
// ===== library types =====

TYPE "UDT_Salidas_RFID"
   STRUCT
      Tag_escribir : Bool;   // Escribir en tag
      Tag_leer : Bool;   // Leer de tag
      Tag_reservado_2 : Bool;   // xBit2
      Tag_reservado_3 : Bool;   // xBit3
      Tag_antena_apagar : Bool;   // Apagar antena
      Tag_reservado_5 : Bool;   // xBit5
      Tag_reservado_6 : Bool;   // xBit6
      Tag_reservado_7 : Bool;   // xBit7
      Reservado_AB5 : Byte;   // byReserved
      Tag_direccion_leer_escribir : Word;   // Direccion de R/W
      Tag_datos_a_escribir : Array[0..27] of Byte;   // Datos a escribir
   END_STRUCT;
END_TYPE

TYPE "UDT_Estado"
   STRUCT
      Modo_auto : Bool;   // Marca Modo
      Modo_manual : Bool;   // Marca Modo
      Ciclo_auto_activo : Bool;   // Marca Modo
      Ciclo_manual_activo : Bool;   // Marca Modo
      Emergencia : Bool;   // Marca Modo
      Rearme_requerido : Bool;   // Marca Modo
      Marcha_permitida : Bool;   // Marca Modo
      Condicion_arranque_auto : Bool;   // Marca Condiciones
      Condicion_arranque_manual : Bool;   // Marca Condiciones
      Estacion_cond_iniciales : Bool;   // Marca Condiciones
      Cinta_habilitada : Bool;   // Marca Condiciones
      Ciclo_manual_terminado : Bool;   // Marca Condiciones
      Rearme_requerido_gestion : Bool;   // Marca Condiciones
      Palet_en_posicion : Bool;   // Marca Cinta
      Palet_en_estacion : Bool;   // Marca Cinta
      Palet_evacuado : Bool;   // Marca Cinta
      Orden_evacuar : Bool;   // Marca Cinta
      Orden_leer : Bool;   // Marca RFID
      Orden_escribir : Bool;   // Marca RFID
      Rfid_lectura_ok : Bool;   // Marca RFID
      Rfid_escritura_ok : Bool;   // Marca RFID
      Rfid_error : Bool;   // Marca RFID
      Rfid_codigo_error : Byte;   // Marca RFID
      App_inicio : Bool;   // Marca App
      App_en_reposo : Bool;   // Marca App
      App_terminada : Bool;   // Marca App
      App_alarma : Bool;
   END_STRUCT;
END_TYPE

TYPE "UDT_Entradas_Basico"
   STRUCT
      Boton_marcha : Bool;   // Botón de marcha
      Boton_paro : Bool;   // Botón de paro (0 activado)
      Selector_modo : Bool;   // Selector Manual/Auto (0 - Manual / 1 - Auto)
      Boton_rearme : Bool;   // Botón de rearme
      Sensor_ind_bien_pos : Bool;   // Palet bien posicionado - Sensor inductivo 0 (Extremo derecho)
      Seta_emergencia : Bool;   // Seta de emergencia
      Sensor_palet_izq : Bool;   // Palet en extremo izquierdo
      Sensor_palet_dch : Bool;   // Palet en extremo derecho
   END_STRUCT;
END_TYPE

TYPE "UDT_Entradas_Stopper"
   STRUCT
      Sensor_ind_0 : Bool;   // Entrada Sensor inductivo 0 (Extremo derecho)
      Sensor_ind_1 : Bool;   // Entrada Sensor inductivo 1
      Sensor_ind_2 : Bool;   // Entrada Sensor inductivo 2
      Sensor_ind_3 : Bool;   // Entrada Sensor inductivo 3 (Extremo izquierdo)
      Reservado_E2_4 : Bool;
      Reservado_E2_5 : Bool;
      Reservado_E2_6 : Bool;
      Sensor_stopper_abajo : Bool;   // Entrada Stopper abajo
   END_STRUCT;
END_TYPE

TYPE "UDT_Salidas_Basico"
   STRUCT
      Led_boton_marcha : Bool;   // Luz del boton de Marcha
      Led_boton_rearme : Bool;   // Luz del boton de Reset
      Led_q1_ciclo_auto : Bool;   // Luz Q1
      Led_q2_emergencia : Bool;   // Luz Q2
      Cinta_dch : Bool;   // Arrancar cinta hacia la derecha
      Cinta_izq : Bool;   // Arrancar cinta hacia la izquierda
      Cinta_velocidad_baja : Bool;   // Establecer velocidad baja
      Bajar_stopper : Bool;   // Bajar cilindro Stopper
   END_STRUCT;
END_TYPE

TYPE "UDT_Entradas_RFID"
   STRUCT
      Tag_datos_escritos : Bool;   // Datos escritos
      Tag_datos_leidos : Bool;   // Datos leidos
      Reservado_E4_2 : Bool;
      Reservado_E4_3 : Bool;
      Tag_antena_apagada : Bool;   // Antena apagada
      Tag_detectado : Bool;   // Tag detectado
      Tag_error : Bool;   // Error
      Tag_proceso_listo : Bool;   // Proceso listo
      Tag_codigo_error : Byte;   // Codigo de error
      Tag_direccion_confirmada : Word;   // Direccion de escritura
      Tag_datos_leidos_escritos : Array[0..27] of Byte;   // Datos
   END_STRUCT;
END_TYPE

FUNCTION_BLOCK "Est_FB_Estacion"   // FB1, SCL
{ S7_Optimized_Access := 'TRUE' }
VERSION : 0.1
   VAR_INPUT
      InBasico : "UDT_Entradas_Basico";
      InRFID : "UDT_Entradas_RFID";
      InStopper : "UDT_Entradas_Stopper";
      Direccion_lectura : Word;
      Direccion_escritura : Word;
      App_en_reposo : Bool;
      App_terminada : Bool;
      App_alarma : Bool;
      App_rearme_requerido : Bool;
      Inhibir_cinta : Bool;
      Mascara_lectura : DWord := 16#0FFFFFFF;
      Mascara_escritura : DWord;
   END_VAR
   VAR_OUTPUT
      App_inicio : Bool;
      Emergencia : Bool;
      Rearme : Bool;
   END_VAR
   VAR_IN_OUT
      OutBasico : "UDT_Salidas_Basico";
      OutRFID : "UDT_Salidas_RFID";
      Imagen_palet : Array[0..27] of Byte;
   END_VAR
   VAR
      Etapa_gestion : Int;
      Etapa_0 : Bool;
      Etapa_1 : Bool;
      Etapa_2 : Bool;
      Etapa_3 : Bool;
      Etapa_4 : Bool;
      Etapa_5 : Bool;
      Estado_Estacion : "UDT_Estado";
      Flanco_rearme : R_TRIG;
      FB2_Modo_Instance : "Est_FB_Modo";
      FB3_Cinta_Instance : "Est_FB_Cinta";
      FB4_RFID_Instance : "Est_FB_RFID";
      Ciclo_manual_acabado : Bool;
   END_VAR
BEGIN
   #Estado_Estacion.App_en_reposo := #App_en_reposo;
   #Estado_Estacion.App_terminada := #App_terminada;
   #Estado_Estacion.App_alarma := #App_alarma;

   //Flanco de rearme
   #Flanco_rearme(CLK := #InBasico.Boton_rearme);

   //Condiciones combinacionales
   //las CI han cambiado ahora que tenemos app
   // Tensión en la máquina (24 Vdc) – No existe señal de PLC.
   // Aire comprimido (6 bar) – No existe señal de PLC.
   // Debe existir un palet correctamente posicionado.
   // El cilindro eje vertical Debe estar en su posición extrema superior.
   // El cilindro eje horizontal Debe estar referenciado.
   // La garra estará en posición de reposo (desctivada/cerrada).
   // No existe estado de emergencia.
   #Estado_Estacion.Estacion_cond_iniciales := NOT #Estado_Estacion.Emergencia AND NOT #InStopper.Sensor_stopper_abajo AND #Estado_Estacion.App_en_reposo
   AND NOT #Estado_Estacion.Rfid_error;

   #Estado_Estacion.Condicion_arranque_auto := #Estado_Estacion.Estacion_cond_iniciales;
   #Estado_Estacion.Condicion_arranque_manual := #Estado_Estacion.Estacion_cond_iniciales AND #Estado_Estacion.Palet_en_estacion;

   #Estado_Estacion.Cinta_habilitada := (#Estado_Estacion.Ciclo_auto_activo OR #Estado_Estacion.Ciclo_manual_activo) AND NOT #Estado_Estacion.Emergencia;

   //llamo a Modo
   #FB2_Modo_Instance(Seta_emergencia := NOT #InBasico.Seta_emergencia,
                      Boton_rearme := #InBasico.Boton_rearme,
                      Boton_marcha := #InBasico.Boton_marcha,
                      Boton_paro := NOT #InBasico.Boton_paro,
                      Selector_automatico := #InBasico.Selector_modo,
                      Condicion_arranque_auto := #Estado_Estacion.Condicion_arranque_auto,
                      Condicion_arranque_manual := #Estado_Estacion.Condicion_arranque_manual,
                      Ciclo_manual_acabado := #Ciclo_manual_acabado,
                      Modo_auto := #Estado_Estacion.Modo_auto,
                      Modo_manual := #Estado_Estacion.Modo_manual,
                      Ciclo_auto_activo := #Estado_Estacion.Ciclo_auto_activo,
                      Ciclo_manual_activo := #Estado_Estacion.Ciclo_manual_activo,
                      Emergencia := #Estado_Estacion.Emergencia,
                      Rearme_requerido := #Estado_Estacion.Rearme_requerido,
                      Marcha_permitida := #Estado_Estacion.Marcha_permitida
   );

   //gestión
   CASE #Etapa_gestion OF
       0:  // ESPERA PALET
           IF (#Estado_Estacion.Ciclo_auto_activo OR #Estado_Estacion.Ciclo_manual_activo) AND #Estado_Estacion.Palet_en_posicion AND NOT #Estado_Estacion.Emergencia THEN
               #Etapa_gestion := 1;
           END_IF;
       1:  // LEER RFID
           IF #Estado_Estacion.Rfid_error THEN
               #Etapa_gestion := 6;
           ELSIF #Estado_Estacion.Rfid_lectura_ok THEN
               #Etapa_gestion := 2;
           END_IF;
       2:  // APLICACION
           IF #Estado_Estacion.App_terminada THEN
               #Etapa_gestion := 3;
           END_IF;
       3:  // ESCRIBIR RFID
           IF #Estado_Estacion.Rfid_error THEN
               #Etapa_gestion := 6;
           ELSIF #Estado_Estacion.Rfid_escritura_ok THEN
               #Etapa_gestion := 4;
           END_IF;
       4:  // EVACUAR
           IF #Estado_Estacion.Palet_evacuado THEN
               #Etapa_gestion := 5;
           END_IF;
       5:  // FIN PALET
           #Etapa_gestion := 0;
       6:  // FALLO RFID
           IF #Flanco_rearme.Q THEN
               #Etapa_gestion := 4;
           END_IF;
       ELSE
           #Etapa_gestion := 0;
   END_CASE;

   //Emergencia
   IF #Estado_Estacion.Emergencia THEN
       #Etapa_gestion := 0;
   END_IF;

   //Ordenes
   #Estado_Estacion.Orden_leer := (#Etapa_gestion = 1);
   #Estado_Estacion.App_inicio := (#Etapa_gestion = 2);
   #Estado_Estacion.Orden_escribir := (#Etapa_gestion = 3);
   #Estado_Estacion.Orden_evacuar := (#Etapa_gestion = 4);
   #Ciclo_manual_acabado := (#Etapa_gestion = 5 OR (#Etapa_gestion = 0 AND NOT #Estado_Estacion.Palet_en_estacion))
   AND #Estado_Estacion.Modo_manual;
   #Estado_Estacion.Rearme_requerido_gestion := (#Etapa_gestion = 6);

   //Cadenas
   #FB3_Cinta_Instance(Cinta_habilitada := #Estado_Estacion.Cinta_habilitada,
                       Orden_evacuar := #Estado_Estacion.Orden_evacuar,
                       Emergencia := #Estado_Estacion.Emergencia,
                       Sensor_palet_izq := #InBasico.Sensor_palet_izq,
                       Sensor_palet_dch := #InBasico.Sensor_palet_dch,
                       Sensor_ind_bien_pos := #InBasico.Sensor_ind_bien_pos,
                       Sensor_stopper_abajo := #InStopper.Sensor_stopper_abajo,
                       Cinta_dch := #OutBasico.Cinta_dch,
                       Bajar_stopper := #OutBasico.Bajar_stopper,
                       Palet_en_posicion := #Estado_Estacion.Palet_en_posicion,
                       Palet_en_estacion := #Estado_Estacion.Palet_en_estacion,
                       Palet_evacuado := #Estado_Estacion.Palet_evacuado
   );

   IF #Inhibir_cinta THEN
       #OutBasico.Cinta_dch := FALSE;
   END_IF;

   #FB4_RFID_Instance(Orden_leer := #Estado_Estacion.Orden_leer,
                      Orden_escribir := #Estado_Estacion.Orden_escribir,
                      Emergencia := #Estado_Estacion.Emergencia,
                      Tag_datos_escritos := #InRFID.Tag_datos_escritos,
                      Tag_datos_leidos := #InRFID.Tag_datos_leidos,
                      Tag_antena_apagada := #InRFID.Tag_antena_apagada,
                      Tag_detectado := #InRFID.Tag_detectado,
                      Tag_error := #InRFID.Tag_error,
                      Tag_proceso_listo := #InRFID.Tag_proceso_listo,
                      Tag_codigo_error := #InRFID.Tag_codigo_error,
                      Tag_direccion_confirmada := #InRFID.Tag_direccion_confirmada,
                      Tag_datos_leidos_escritos := #InRFID.Tag_datos_leidos_escritos,
                      Mascara_lectura:=#Mascara_lectura,
                      Mascara_escritura:=#Mascara_escritura,
                      Tag_escribir := #OutRFID.Tag_escribir,
                      Tag_leer := #OutRFID.Tag_leer,
                      Tag_antena_apagar := #OutRFID.Tag_antena_apagar,
                      Tag_direccion_leer_escribir := #OutRFID.Tag_direccion_leer_escribir,
                      Tag_datos_a_escribir := #OutRFID.Tag_datos_a_escribir,
                      Rfid_lectura_ok := #Estado_Estacion.Rfid_lectura_ok,
                      Rfid_escritura_ok := #Estado_Estacion.Rfid_escritura_ok,
                      Rfid_error := #Estado_Estacion.Rfid_error,
                      Rfid_codigo_error := #Estado_Estacion.Rfid_codigo_error,
                      Imagen:=#Imagen_palet,
                      Direccion_escritura:=#Direccion_escritura,
                      Direccion_lectura:=#Direccion_lectura);

   #App_inicio := #Estado_Estacion.App_inicio;
   #Emergencia := #Estado_Estacion.Emergencia;
   #Rearme := #Flanco_rearme.Q;

   //Luces del panel y salidas sin uso
   #OutBasico.Led_boton_marcha := #Estado_Estacion.Marcha_permitida;
   #OutBasico.Led_boton_rearme := #Estado_Estacion.Rearme_requerido OR #Estado_Estacion.Rearme_requerido_gestion OR #App_rearme_requerido;
   #OutBasico.Led_q1_ciclo_auto := #Estado_Estacion.Ciclo_auto_activo;
   #OutBasico.Led_q2_emergencia := #Estado_Estacion.Emergencia OR (#Estado_Estacion.App_alarma);// AND "Clock_1Hz");
   #OutBasico.Cinta_izq := FALSE;
   #OutBasico.Cinta_velocidad_baja := FALSE;
END_FUNCTION_BLOCK

FUNCTION_BLOCK "Est_FB_Modo"   // FB2, SCL
{ S7_Optimized_Access := 'TRUE' }
VERSION : 0.1
   VAR_INPUT
      Seta_emergencia : Bool;
      Boton_rearme : Bool;
      Boton_marcha : Bool;
      Boton_paro : Bool;
      Selector_automatico : Bool;
      Condicion_arranque_auto : Bool;
      Condicion_arranque_manual : Bool;
      Ciclo_manual_acabado : Bool;
   END_VAR
   VAR_IN_OUT
      Modo_auto : Bool;
      Modo_manual : Bool;
      Ciclo_auto_activo : Bool;
      Ciclo_manual_activo : Bool;
      Emergencia : Bool;
      Rearme_requerido : Bool;
      Marcha_permitida : Bool;
   END_VAR
   VAR
      Etapa_emergencia : Int := 10;
      Etapa_modo : Int := 20;
      Etapa_ciclo : Int := 30;
      Flanco_marcha : R_TRIG;
      Flanco_rearme : R_TRIG;
   END_VAR
BEGIN
   #Modo_auto := FALSE;
   #Modo_manual := FALSE;
   #Ciclo_auto_activo := FALSE;
   #Ciclo_manual_activo := FALSE;
   #Emergencia := FALSE;
   #Rearme_requerido := FALSE;
   #Marcha_permitida := FALSE;

   #Flanco_marcha(CLK:=#Boton_marcha);
   #Flanco_rearme(CLK:=#Boton_rearme);

   CASE #Etapa_emergencia OF
       10:  //NORMAL
           IF #Seta_emergencia THEN
               #Etapa_emergencia := 11;
           END_IF;
           ;
       11:  //EMERGENCIA
           #Emergencia := TRUE;
           #Rearme_requerido := TRUE;
           IF #Flanco_rearme.Q AND NOT #Seta_emergencia THEN
               #Etapa_emergencia := 10;
           END_IF;
           ;
       ELSE
           #Etapa_emergencia := 11;
           ;
   END_CASE;

   CASE #Etapa_modo OF
       20:  // MANUAL
           #Modo_manual := TRUE;
           IF #Selector_automatico THEN
               #Etapa_modo := 21;
           END_IF;
           ;
       21:  // AUTOMATICO
           #Modo_auto := TRUE;
           IF NOT #Selector_automatico THEN
               #Etapa_modo := 20;
           END_IF;
           ;
       ELSE
           #Etapa_modo := 20;
           #Etapa_emergencia := 11;
           ;
   END_CASE;

   CASE #Etapa_ciclo OF
       30:  // REPOSO
           IF NOT #Emergencia AND ((#Modo_auto AND #Condicion_arranque_auto) OR (#Modo_manual AND #Condicion_arranque_manual)) THEN
               #Marcha_permitida := TRUE;
           END_IF;

           IF #Marcha_permitida AND #Flanco_marcha.Q AND #Modo_auto THEN
               #Etapa_ciclo := 31;
           ELSIF #Marcha_permitida AND #Flanco_marcha.Q AND #Modo_manual THEN
               #Etapa_ciclo := 32;
           END_IF;
           ;
       31:  // AUTOMATICO ACTIVO
           #Ciclo_auto_activo := TRUE;
           IF #Boton_paro OR #Emergencia OR NOT #Modo_auto THEN
               #Etapa_ciclo := 30;
           END_IF;
           ;
       32:  //MANUAL ACTIVO
           #Ciclo_manual_activo := TRUE;
           IF #Boton_paro OR #Emergencia OR NOT #Modo_manual OR #Ciclo_manual_acabado THEN
               #Etapa_ciclo := 30;
           END_IF;
           ;
       ELSE
           #Etapa_ciclo := 30;
           #Etapa_emergencia := 11;
           ;
   END_CASE;
END_FUNCTION_BLOCK

FUNCTION_BLOCK "Est_FB_Cinta"   // FB3, SCL
{ S7_Optimized_Access := 'TRUE' }
VERSION : 0.1
   VAR_INPUT
      Emergencia : Bool;   // De modo
      Cinta_habilitada : Bool;   // ciclo activo y estación en condiciones iniciales
      Orden_evacuar : Bool;   // la aplicación ya terminó y el RFID está escrito
      Sensor_palet_izq : Bool;   // Extremos de la cinta
      Sensor_palet_dch : Bool;   // Extremos de la cinta
      Sensor_ind_bien_pos : Bool;   // Palet apoyado en el stopper
      Sensor_stopper_abajo : Bool;   // Confirmación del stopper
   END_VAR
   VAR_IN_OUT
      Cinta_dch : Bool;   // Actuadores
      Bajar_stopper : Bool;   // Actuadores
      Palet_en_posicion : Bool;   // Hay palet listo para trabajar
      Palet_en_estacion : Bool;   // Sensor_palet_izq + Sensor_palet_dch + Sensor_ind_bien_pos, para Condicion_arranque_manual
      Palet_evacuado : Bool;   // activa Ciclo_manual_terminado
   END_VAR
   VAR
      Etapa_cinta : Int;   // nuemero de etapa
      Etapa_2 : Bool;   // estamos en la 2
      Timer_etapa2 : TON_TIME;   // timer de la 2
      Flanco_subida_sensor_palet_dch : R_TRIG;   // flanco subida del sensor
      Flanco_bajada_sensor_palet_dch : F_TRIG;   // flanco bajada del sensor
      Palets_en_cinta : Int;
      Flanco_subida_sensor_palet_izq : R_TRIG;
      Timer_Stopper_Etapa5 : TON_TIME;
      Timer_avance : TON_TIME;
   END_VAR
BEGIN

   #Cinta_dch := FALSE;
   #Palet_en_posicion := FALSE;
   #Palet_en_estacion := FALSE;
   #Etapa_2 := FALSE;
   #Palet_evacuado := FALSE;

   #Flanco_subida_sensor_palet_dch(CLK := #Sensor_palet_dch);
   #Flanco_bajada_sensor_palet_dch(CLK := #Sensor_palet_dch);
   #Flanco_subida_sensor_palet_izq(CLK := #Sensor_palet_izq);
   #Timer_Stopper_Etapa5(IN := #Etapa_cinta = 5,
                         PT := T#400ms);
   #Timer_avance(IN := #Etapa_cinta = 1 OR #Etapa_cinta = 6, PT := T#10s);



   IF #Etapa_cinta = 2 THEN
       #Etapa_2 := TRUE;
   END_IF;

   #Timer_etapa2(IN := #Etapa_2,
                 PT := T#300ms);

   IF #Flanco_subida_sensor_palet_izq.Q THEN
       #Palets_en_cinta := #Palets_en_cinta + 1;
   END_IF;
   IF #Flanco_bajada_sensor_palet_dch.Q AND #Palets_en_cinta > 0 THEN
       #Palets_en_cinta := #Palets_en_cinta - 1;
   END_IF;

   IF #Sensor_ind_bien_pos AND #Palets_en_cinta = 0 THEN
       #Palets_en_cinta := 1;
   END_IF;

   CASE #Etapa_cinta OF
       0:  // PARADA
           #Cinta_dch := FALSE;
           #Bajar_stopper := FALSE;
           IF #Cinta_habilitada AND (#Sensor_palet_izq OR #Palets_en_cinta > 0) AND NOT #Sensor_ind_bien_pos THEN
               #Etapa_cinta := 1;
           ELSIF #Cinta_habilitada AND #Sensor_ind_bien_pos THEN
               #Etapa_cinta := 3;
           END_IF;
       1:  //AVANCE
           #Cinta_dch := TRUE;
           IF #Sensor_ind_bien_pos THEN
               #Etapa_cinta := 3;
           ELSIF #Timer_avance.Q THEN   // no llega ningun palet: el contador estaba descuadrado
               #Palets_en_cinta := 0;
               #Etapa_cinta := 0;
           END_IF;
       2:  //ASENTAR
           #Cinta_dch := TRUE;
           IF #Timer_etapa2.Q THEN
               #Etapa_cinta := 3;
           END_IF;
       3:  //PALET EN POSICION
           #Palet_en_posicion := TRUE;
           IF #Orden_evacuar THEN
               #Etapa_cinta := 4;
           END_IF;
       4:  //LIBERAR
           #Bajar_stopper := TRUE;
           IF NOT #Sensor_stopper_abajo THEN
               #Etapa_cinta := 5;
           END_IF;
       5:  //SACAR
           #Bajar_stopper := TRUE;
           #Cinta_dch := TRUE;
           IF #Timer_Stopper_Etapa5.Q OR #Flanco_subida_sensor_palet_dch.Q THEN
               #Etapa_cinta := 6;
               ;
           END_IF;
       6: //SALIR
           #Bajar_stopper := FALSE;
           #Cinta_dch := TRUE;
           IF #Flanco_bajada_sensor_palet_dch.Q THEN
               #Etapa_cinta := 7;
               ;
           ELSIF #Timer_avance.Q THEN   // el palet no pasa por el sensor (retirado a mano): no dejar la cinta en marcha
               #Palets_en_cinta := 0;
               #Etapa_cinta := 7;
           END_IF;
       7: //TERMINAR
           #Palet_evacuado := TRUE;
           #Etapa_cinta := 0;
       ELSE  // Statement section ELSE
           #Etapa_cinta := 0;
           ;
   END_CASE;

   #Palet_en_estacion := #Sensor_palet_dch OR #Sensor_palet_izq OR #Sensor_ind_bien_pos OR (#Palets_en_cinta > 0) OR #Etapa_cinta = 1;

   IF #Emergencia THEN
       #Etapa_cinta := 0;
       #Cinta_dch := FALSE;
       #Bajar_stopper := FALSE;
       #Palets_en_cinta := 0;   // el operario retira los palets en la emergencia
   END_IF;
END_FUNCTION_BLOCK

FUNCTION_BLOCK "Est_FB_RFID"   // FB4, SCL
{ S7_Optimized_Access := 'TRUE' }
VERSION : 0.1
   VAR_INPUT
      Emergencia : Bool;
      Orden_escribir : Bool;
      Orden_leer : Bool;
      Tag_datos_escritos : Bool;
      Tag_datos_leidos : Bool;
      Tag_antena_apagada : Bool;
      Tag_detectado : Bool;
      Tag_error : Bool;
      Tag_proceso_listo : Bool;
      Tag_codigo_error : Byte;
      Tag_direccion_confirmada : Word;
      Tag_datos_leidos_escritos : Array[0..27] of Byte;
      Direccion_lectura : Word;
      Direccion_escritura : Word;
      Mascara_lectura : DWord;
      Mascara_escritura : DWord;
   END_VAR
   VAR_IN_OUT
      Tag_escribir : Bool;
      Tag_leer : Bool;
      Tag_antena_apagar : Bool;
      Tag_direccion_leer_escribir : Word;
      Tag_datos_a_escribir : Array[0..27] of Byte;
      Rfid_lectura_ok : Bool;
      Rfid_escritura_ok : Bool;
      Rfid_error : Bool;
      Rfid_codigo_error : Byte;
      Imagen : Array[0..27] of Byte;
   END_VAR
   VAR
      T_Rfid : TON_TIME;
      Etapa_rfid : Int;
      Etapa_1 : Bool;
      Etapa_3 : Bool;
      Etapa_4 : Bool;
      Rfid_ocupado : Bool;
      Imagen_leida : Array[0..27] of Byte;
   END_VAR
   VAR_TEMP
      i : Int;
   END_VAR
BEGIN
   //PARA EL DANI DEL FUTURO
   //que vaya leyendo los codigos rfid por si me vienen dos palets juntos
   //y que los meta en una cola para luego leerlos y escribirlos por orden?
   //      - no lo voy a hacer porque creo que esto solo es un problema en el simulador
   //      - pero gracias por la idea dani del pasado
   //---------------------------------------------------------------------------
   #Tag_escribir := FALSE;
   #Tag_leer := FALSE;
   #Tag_antena_apagar := TRUE;
   #Rfid_lectura_ok := FALSE;
   #Rfid_escritura_ok := FALSE;
   #Rfid_error := FALSE;
   #Etapa_1 := FALSE;
   #Etapa_3 := FALSE;
   #Etapa_4 := FALSE;

   CASE #Etapa_rfid OF
       0:  // REPOSO
           #Tag_antena_apagar := TRUE;
           #Tag_leer := FALSE;
           #Tag_escribir := FALSE;
           IF (#Orden_leer OR #Orden_escribir) AND NOT #Emergencia THEN
               #Etapa_rfid := 1;
               ;
           END_IF;
       1:  // ENERGIZAR
           #Tag_antena_apagar := FALSE;
           #Etapa_1 := TRUE;
           IF #Tag_error OR #T_Rfid.Q THEN
               #Etapa_rfid := 8;
           ELSIF NOT #Tag_antena_apagada AND #Tag_detectado AND #Tag_proceso_listo AND NOT #Tag_error THEN
               #Etapa_rfid := 2;
           END_IF;
           ;
       2:  // LISTO
           #Tag_antena_apagar := FALSE;
           #Rfid_ocupado := FALSE;
           IF #Orden_leer AND NOT #Orden_escribir THEN
               #Etapa_rfid := 3;
           ELSIF NOT #Orden_leer AND #Orden_escribir THEN
               #Etapa_rfid := 4;
           END_IF;
           ;
       3:  // LEER
           #Tag_antena_apagar := FALSE;
           #Etapa_3 := TRUE;
           // "leido" es el eco de la orden: el dato solo vale cuando "listo" baja y vuelve a subir
           IF NOT #Tag_proceso_listo THEN
               #Rfid_ocupado := TRUE;
           END_IF;
           #Tag_leer := TRUE;
           #Tag_direccion_leer_escribir := #Direccion_lectura;
           IF #Tag_error OR #T_Rfid.Q THEN
               #Etapa_rfid := 8;
           ELSIF #Rfid_ocupado AND #Tag_datos_leidos AND #Tag_proceso_listo AND #Tag_direccion_confirmada = #Direccion_lectura THEN
               #Imagen_leida := #Tag_datos_leidos_escritos;   // copia completa se usa al escribir
               FOR #i := 0 TO 27 DO
                   IF (SHR(IN := #Mascara_lectura, N := #i) AND 16#1) <> 16#0 THEN
                       #Imagen[#i] := #Tag_datos_leidos_escritos[#i];
                   ELSE
                       #Imagen[#i] := 0;   // lo que no es de esta estacion no pasa a la app
                   END_IF;
               END_FOR;
               #Etapa_rfid := 5;
           END_IF;
           ;
       4:  // ESCRIBIR
           #Tag_antena_apagar := FALSE;
           #Etapa_4 := TRUE;
           IF NOT #Tag_proceso_listo THEN
               #Rfid_ocupado := TRUE;
           END_IF;
           #Tag_escribir := TRUE;
           #Tag_direccion_leer_escribir := #Direccion_escritura;
           FOR #i := 0 TO 27 DO
               IF (SHR(IN := #Mascara_escritura, N := #i) AND 16#1) <> 16#0 THEN
                   #Tag_datos_a_escribir[#i] := #Imagen[#i];       // byte de esta estacion
               ELSE
                   #Tag_datos_a_escribir[#i] := #Imagen_leida[#i]; // byte ajeno: se devuelve como estaba
               END_IF;
           END_FOR;
           IF #Tag_error OR #T_Rfid.Q THEN
               #Etapa_rfid := 8;
           ELSIF #Rfid_ocupado AND #Tag_datos_escritos AND #Tag_proceso_listo AND #Tag_direccion_confirmada = #Direccion_escritura THEN
               #Etapa_rfid := 6;
           END_IF;
           ;
       5:  // LEIDO
           #Tag_antena_apagar := FALSE;
           #Rfid_lectura_ok := TRUE;
           IF NOT #Orden_leer THEN
               #Etapa_rfid := 0;
           END_IF;
           ;
       6:  // ESCRITO 
           #Tag_antena_apagar := FALSE;
           #Rfid_escritura_ok := TRUE;
           IF NOT #Orden_escribir THEN
               #Etapa_rfid := 0;
           END_IF;
           ;
       8:  // ERROR RFID
           #Rfid_error := TRUE;
           #Rfid_codigo_error := #Tag_codigo_error;
           #Tag_antena_apagar := TRUE;
           #Tag_leer := FALSE;
           #Tag_escribir := FALSE;
           IF NOT #Orden_escribir AND NOT #Orden_leer THEN   // CIROS no da "antena apagada" (iAntenaOFF sin conectar)
               #Etapa_rfid := 0;
           END_IF;
           ;
       ELSE  // Statement section ELSE
           #Etapa_rfid := 0;
           ;
   END_CASE;

   #T_Rfid(IN := #Etapa_1 OR #Etapa_3 OR #Etapa_4,
           PT := T#5s);

   IF #Emergencia THEN
       #Etapa_rfid := 0;
       #Tag_antena_apagar := TRUE;
       #Tag_escribir := FALSE;
       #Tag_leer := FALSE;
       #Rfid_lectura_ok := FALSE;
       #Rfid_escritura_ok := FALSE;
       #Rfid_error := FALSE;
   END_IF;
END_FUNCTION_BLOCK

// ===== library: MasterCopy "Main" =====

ORGANIZATION_BLOCK "Main"   // OB1, LAD, ProgramCycle
TITLE = "Main Program Sweep (Cycle)"
{ S7_Optimized_Access := 'TRUE' }
VERSION : 0.1
   VAR_INPUT
      Initial_Call : Bool;   // Initial call of this OB
      Remanence : Bool;   // =True, if remanent data are available
   END_VAR
BEGIN

REGION Network 1: Llamada al gestor
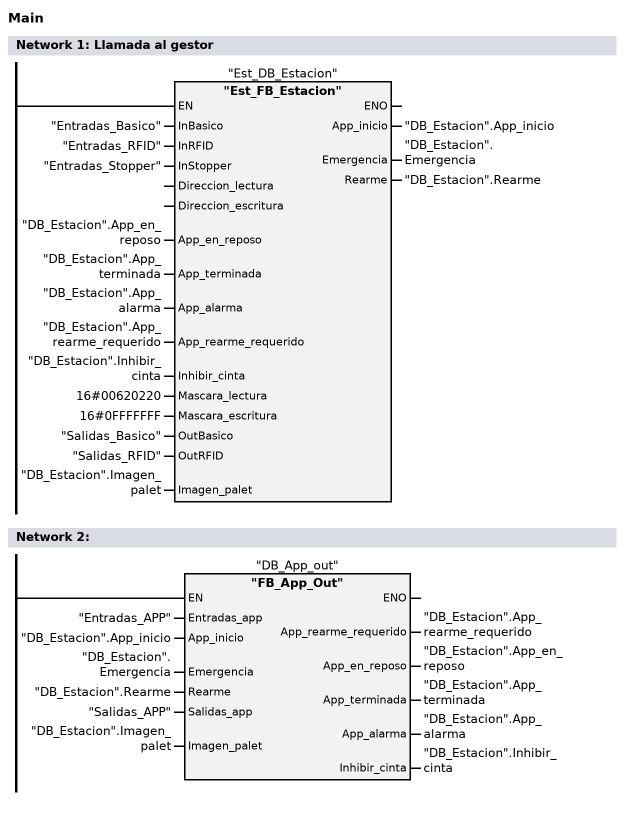
   RUNG wire#powerrail
      "Est_DB_Estacion"(InBasico := "Entradas_Basico", InRFID := "Entradas_RFID", InStopper := "Entradas_Stopper", Direccion_lectura :=, Direccion_escritura :=, App_en_reposo := "DB_Estacion".App_en_reposo, App_terminada := "DB_Estacion".App_terminada, App_alarma := "DB_Estacion".App_alarma, App_rearme_requerido := "DB_Estacion".App_rearme_requerido, Inhibir_cinta := "DB_Estacion".Inhibir_cinta, Mascara_lectura := 16#00620220, Mascara_escritura := 16#0FFFFFFF, OutBasico := "Salidas_Basico", OutRFID := "Salidas_RFID", Imagen_palet := "DB_Estacion".Imagen_palet, App_inicio => "DB_Estacion".App_inicio, Emergencia => "DB_Estacion".Emergencia, Rearme => "DB_Estacion".Rearme)
   END_RUNG
   // the same network as SCL:
   "Est_DB_Estacion"(InBasico := "Entradas_Basico",   // "Est_FB_Estacion"
                     InRFID := "Entradas_RFID",
                     InStopper := "Entradas_Stopper",
                     App_en_reposo := "DB_Estacion".App_en_reposo,
                     App_terminada := "DB_Estacion".App_terminada,
                     App_alarma := "DB_Estacion".App_alarma,
                     App_rearme_requerido := "DB_Estacion".App_rearme_requerido,
                     Inhibir_cinta := "DB_Estacion".Inhibir_cinta,
                     Mascara_lectura := 16#00620220,
                     Mascara_escritura := 16#0FFFFFFF,
                     OutBasico := "Salidas_Basico",
                     OutRFID := "Salidas_RFID",
                     Imagen_palet := "DB_Estacion".Imagen_palet,
                     App_inicio => "DB_Estacion".App_inicio,
                     Emergencia => "DB_Estacion".Emergencia,
                     Rearme => "DB_Estacion".Rearme);
END_REGION

REGION Network 2
   RUNG wire#powerrail
      "DB_App_out"(Entradas_app := "Entradas_APP", App_inicio := "DB_Estacion".App_inicio, Emergencia := "DB_Estacion".Emergencia, Rearme := "DB_Estacion".Rearme, Salidas_app := "Salidas_APP", Imagen_palet := "DB_Estacion".Imagen_palet, App_rearme_requerido => "DB_Estacion".App_rearme_requerido, App_en_reposo => "DB_Estacion".App_en_reposo, App_terminada => "DB_Estacion".App_terminada, App_alarma => "DB_Estacion".App_alarma, Inhibir_cinta => "DB_Estacion".Inhibir_cinta)
   END_RUNG
   // the same network as SCL:
   "DB_App_out"(Entradas_app := "Entradas_APP",   // "FB_App_Out"
                App_inicio := "DB_Estacion".App_inicio,
                Emergencia := "DB_Estacion".Emergencia,
                Rearme := "DB_Estacion".Rearme,
                Salidas_app := "Salidas_APP",
                Imagen_palet := "DB_Estacion".Imagen_palet,
                App_rearme_requerido => "DB_Estacion".App_rearme_requerido,
                App_en_reposo => "DB_Estacion".App_en_reposo,
                App_terminada => "DB_Estacion".App_terminada,
                App_alarma => "DB_Estacion".App_alarma,
                Inhibir_cinta => "DB_Estacion".Inhibir_cinta);
END_REGION
END_ORGANIZATION_BLOCK

// ===== library: MasterCopy "DB_Estacion" =====

DATA_BLOCK "DB_Estacion"   // DB2
{ S7_Optimized_Access := 'TRUE' }
VERSION : 0.1
   VAR
      Imagen_palet : Array[0..27] of Byte;
      App_inicio : Bool;
      App_en_reposo : Bool;
      App_terminada : Bool;
      App_alarma : Bool;
      App_rearme_requerido : Bool;
      Inhibir_cinta : Bool;
      Emergencia : Bool;
      Rearme : Bool;
   END_VAR
BEGIN
END_DATA_BLOCK

// ===== library: MasterCopy "FB_App_Out" =====

FUNCTION_BLOCK "FB_App_Out"   // FB5, SCL
{ S7_Optimized_Access := 'TRUE' }
VERSION : 0.1
   VAR_INPUT
      Entradas_app : "UDT_Entradas_APP";
      App_inicio : Bool;
      Emergencia : Bool;
      Rearme : Bool;
   END_VAR
   VAR_OUTPUT
      App_rearme_requerido : Bool;
      App_en_reposo : Bool;
      App_terminada : Bool;
      App_alarma : Bool;
      Inhibir_cinta : Bool;
   END_VAR
   VAR_IN_OUT
      Salidas_app : "UDT_Salidas_APP";
      Imagen_palet : Array[0..27] of Byte;
   END_VAR
   VAR
      Cond_conf : Bool;
      Cond_almacen : Bool;
      Etapa_app : Int;
      Etapa_previa : Int;
      Posicion_objetivo : Int;
      Almacen_destino : Int;
      Start_enviado : Bool;
      Pieza_en_garra : Bool;
      Parpadeo : Bool;
      Emergencia_previa : Bool;
      Recuperando : Bool;
      Timer_arranque : TON_TIME;
      Timer_conf : TON_TIME;
      Timer_almacen : TON_TIME;
      Timer_parpadeo : TON_TIME;
      Timer_freno : TON_TIME;
   END_VAR
   VAR_TEMP
      i : Int;
   END_VAR
   VAR CONSTANT
      IDX_CALIDAD : Int := 5;
      IDX_DESTINO : Int := 17;
   END_VAR
BEGIN
   #App_en_reposo := FALSE;
   #App_terminada := FALSE;
   #Cond_conf := FALSE;
   #Cond_almacen := FALSE;
   #Salidas_app.Bajar_cilindro := FALSE;
   #Salidas_app.Subir_cilindro := FALSE;
   #Salidas_app.Abrir_freno := FALSE;     // FALSE = freno puesto
   #Salidas_app.Abrir_garra := FALSE;     // FALSE = garra cerrada
   #Salidas_app.Iniciar_mov_driver_motor := FALSE;
   #Salidas_app.Activar_driver_motor := NOT #Emergencia;

   CASE #Etapa_app OF
       0:  // REPOSO
           #App_en_reposo := #Entradas_app.Eje_z_arriba AND NOT #Entradas_app.Gripper_abierto
           AND #Entradas_app.Eje_referenciado AND NOT #Pieza_en_garra;
           IF #Pieza_en_garra AND #Entradas_app.Eje_z_arriba AND #Entradas_app.Eje_referenciado THEN
               #Almacen_destino := 1;          // tapa de una emergencia: al almacen de erroneas
               #Posicion_objetivo := 3;
               #Recuperando := TRUE;
               #Etapa_app := 7;
           ELSIF #App_inicio AND #App_en_reposo THEN
               IF #Imagen_palet[#IDX_DESTINO] = 1 OR #Imagen_palet[#IDX_DESTINO] = 2 THEN
                   #Almacen_destino := BYTE_TO_INT(#Imagen_palet[#IDX_DESTINO]);   // forzado por receta: 1 izq, 2 dcha
               ELSIF #Imagen_palet[#IDX_CALIDAD] = 1 THEN
                   #Almacen_destino := 2;   // calidad OK -> derecho
               ELSE
                   #Almacen_destino := 1;   // NOK o sin evaluar -> izquierdo
               END_IF;
               #Posicion_objetivo := 3;        // 3 = centro
               #Etapa_app := 1;
           ELSIF NOT #App_en_reposo THEN
               #Etapa_app := 20;               // recolocar / referenciar
           END_IF;

       1, 7, 11:  // ORDEN DE MOVIMIENTO (flanco de START, MC cae = arranca)
           IF NOT #Start_enviado THEN
               #Start_enviado := #Entradas_app.Eje_z_arriba AND #Entradas_app.Ready AND #Entradas_app.Motion_complete;
           ELSE
               #Salidas_app.Iniciar_mov_driver_motor := #Entradas_app.Eje_z_arriba;
               IF NOT #Entradas_app.Motion_complete OR #Timer_arranque.Q THEN
                   #Start_enviado := FALSE;
                   #Etapa_app := #Etapa_app + 1;
               END_IF;
           END_IF;
           IF #Etapa_app = 11 OR #Etapa_app = 12 THEN
               #Salidas_app.Abrir_garra := TRUE;   // al volver, la garra sigue abierta
           END_IF;

       2, 8, 12, 22:  // ESPERAR FIN DE MOVIMIENTO (START a 0, MC sube = posicion alcanzada)
           IF #Etapa_app = 12 THEN
               #Salidas_app.Abrir_garra := TRUE;
           END_IF;
           IF #Entradas_app.Motion_complete THEN
               IF #Etapa_app = 8 AND #Posicion_objetivo = 3 THEN
                   #Etapa_app := 9;
               ELSIF #Etapa_app = 8 THEN
                   #Etapa_app := 10;
               ELSE
                   #Etapa_app := #Etapa_app + 1;
               END_IF;
           END_IF;

       3:  // ABRIR GARRA
           #Salidas_app.Abrir_garra := TRUE;
           IF #Entradas_app.Gripper_abierto THEN
               #Etapa_app := 4;
           END_IF;

       4:  // BAJAR Z (primero se abre el freno, la bajada entra un ciclo despues)
           #Salidas_app.Abrir_garra := TRUE;
           #Salidas_app.Abrir_freno := TRUE;
           #Salidas_app.Bajar_cilindro := #Etapa_app = #Etapa_previa;
           #Cond_conf := #Entradas_app.Eje_z_abajo;
           IF #Timer_conf.Q THEN
               #Etapa_app := 5;
           END_IF;

       5:  // CERRAR GARRA
           #Salidas_app.Abrir_freno := TRUE;
           #Salidas_app.Bajar_cilindro := TRUE;
           #Cond_conf := NOT #Entradas_app.Gripper_abierto;
           IF #Timer_conf.Q THEN
               #Pieza_en_garra := TRUE;
               #Etapa_app := 6;
           END_IF;

       6:  // SUBIR Z
           #Salidas_app.Abrir_freno := TRUE;
           #Salidas_app.Subir_cilindro := TRUE;
           #Cond_conf := #Entradas_app.Eje_z_arriba;
           IF #Timer_conf.Q THEN
               #Etapa_app := 9;
           END_IF;

       9:  // ESPERAR ALMACEN LIBRE
           #Cond_almacen := (#Almacen_destino = 1 AND #Entradas_app.Almacen_izq_lleno)
           OR (#Almacen_destino = 2 AND #Entradas_app.Almacen_dch_lleno);
           IF NOT #Cond_almacen THEN
               #Posicion_objetivo := #Almacen_destino;
               #Etapa_app := 7;
           END_IF;

       10: // SOLTAR PIEZA
           #Salidas_app.Abrir_garra := TRUE;
           #Cond_conf := #Entradas_app.Gripper_abierto;
           IF #Timer_conf.Q THEN
               #Pieza_en_garra := FALSE;
               #Posicion_objetivo := 3;
               #Etapa_app := 11;
           END_IF;

       13: // CERRAR GARRA
           #Cond_conf := NOT #Entradas_app.Gripper_abierto;
           IF #Timer_conf.Q AND #Recuperando THEN
               #Recuperando := FALSE;
               #Etapa_app := 0;                // sin App_terminada: no habia ciclo de gestion
           ELSIF #Timer_conf.Q THEN
               #Etapa_app := 14;
           END_IF;

       14: // FIN
           FOR #i := 0 TO 27 DO
               #Imagen_palet[#i] := 0;   // la tabla pide dejar el palet limpio para la siguiente vuelta
           END_FOR;
           #App_terminada := TRUE;
           IF NOT #App_inicio THEN
               #Etapa_app := 0;
           END_IF;

       20: // RECOLOCAR: subir Z con garra cerrada (primero aire, luego freno; si Z ya esta arriba el freno no se abre)
           #Salidas_app.Abrir_freno := #Timer_freno.Q;
           #Salidas_app.Subir_cilindro := TRUE;
           #Cond_conf := #Entradas_app.Eje_z_arriba AND NOT #Entradas_app.Gripper_abierto;
           IF #Timer_conf.Q THEN
               IF #Entradas_app.Eje_referenciado THEN
                   #Etapa_app := 0;
               ELSE
                   #Posicion_objetivo := 0;    // 00 = referenciar
                   #Etapa_app := 21;
               END_IF;
           END_IF;

       21: // REFERENCIAR: START con bits 00 sin esperar Ready/MC (Ready no sube hasta estar referenciado)
           #Salidas_app.Iniciar_mov_driver_motor := #Entradas_app.Eje_z_arriba AND #Etapa_app = #Etapa_previa;
           IF #Entradas_app.Eje_referenciado THEN
               #Etapa_app := 22;
           END_IF;

       23: // FIN REFERENCIADO
           #Etapa_app := 0;

       30: // ESPERA REARME (arranque y tras emergencia): nada se mueve
           IF (#Rearme OR #Emergencia_previa) AND NOT #Emergencia THEN
               #Etapa_app := 20;
           END_IF;

       ELSE
           #Etapa_app := 20;
   END_CASE;

   //Bits de posicion del driver (Bit1 Bit0): 00 ref, 01 izq, 10 dch, 11 centro
   #Salidas_app.Bit_pos_0 := (#Posicion_objetivo = 1) OR (#Posicion_objetivo = 3);
   #Salidas_app.Bit_pos_1 := (#Posicion_objetivo = 2) OR (#Posicion_objetivo = 3);

   //Temporizadores (Timer_conf se resetea en cada cambio de etapa)
   #Timer_arranque(IN := #Start_enviado,
                   PT := T#500ms);
   #Timer_conf(IN := #Cond_conf AND #Etapa_app = #Etapa_previa,
               PT := T#300ms);
   #Timer_almacen(IN := #Cond_almacen,
                  PT := T#10s);
   #Timer_parpadeo(IN := #Timer_almacen.Q AND NOT #Timer_parpadeo.Q,
                   PT := T#500ms);
   #Timer_freno(IN := #Etapa_app = 20 AND #Etapa_previa = 20,
                PT := T#500ms);
   IF #Timer_parpadeo.Q THEN
       #Parpadeo := NOT #Parpadeo;
   END_IF;
   #App_alarma := #Timer_almacen.Q AND #Parpadeo;
   #Etapa_previa := #Etapa_app;
   #Emergencia_previa := #Emergencia;

   //X no se mueve si Z no esta arriba
   IF NOT #Entradas_app.Eje_z_arriba THEN
       #Salidas_app.Iniciar_mov_driver_motor := FALSE;
   END_IF;

   //Emergencia
   IF #Emergencia THEN
       IF #Entradas_app.Eje_z_abajo AND (#Etapa_app = 4 OR #Etapa_app = 5) THEN
           #Pieza_en_garra := TRUE;    // la garra se cierra al quitar la salida y atrapa la tapa
       END_IF;
       #Recuperando := FALSE;
       #Etapa_app := 30;
       #Start_enviado := FALSE;
       #Salidas_app.Bajar_cilindro := FALSE;
       #Salidas_app.Subir_cilindro := FALSE;
       #Salidas_app.Abrir_freno := FALSE;
       #Salidas_app.Abrir_garra := FALSE;
       #Salidas_app.Iniciar_mov_driver_motor := FALSE;
       #Salidas_app.Activar_driver_motor := FALSE;
       #Salidas_app.Bit_pos_0 := FALSE;
       #Salidas_app.Bit_pos_1 := FALSE;
   END_IF;

   #Inhibir_cinta := NOT #Entradas_app.Eje_z_arriba; //la cinta no se mueve con Z abajo
   #App_rearme_requerido := #Etapa_app = 30;
END_FUNCTION_BLOCK

// ===== library: MasterCopy "DB_App_out" =====

DATA_BLOCK "DB_App_out"   // DB3
{ S7_Optimized_Access := 'TRUE' }
VERSION : 0.1
// stored: InstanceOfName FB_App_Out
"FB_App_Out"
BEGIN
END_DATA_BLOCK

// ===== library: MasterCopy "UDT_Entradas_APP" =====

TYPE "UDT_Entradas_APP"
   STRUCT
      Eje_z_arriba : Bool;
      Eje_z_abajo : Bool;
      Gripper_abierto : Bool;
      Almacen_izq_lleno : Bool;
      Almacen_dch_lleno : Bool;
      Eje_referenciado : Bool;
      Motion_complete : Bool;
      Ready : Bool;
   END_STRUCT;
END_TYPE

// ===== library: MasterCopy "UDT_Salidas_APP" =====

TYPE "UDT_Salidas_APP"
   STRUCT
      Subir_cilindro : Bool;
      Bajar_cilindro : Bool;
      Abrir_freno : Bool;
      Abrir_garra : Bool;
      Activar_driver_motor : Bool;
      Bit_pos_0 : Bool;
      Bit_pos_1 : Bool;
      Iniciar_mov_driver_motor : Bool;
   END_STRUCT;
END_TYPE

// ===== library: MasterCopy "Tabla de variables estándar" =====

VAR_GLOBAL   // PLC tag table "Tabla de variables estándar"
   "Entradas_APP" AT %E0.0 : "UDT_Entradas_APP";
   "Entradas_Basico" AT %E1.0 : "UDT_Entradas_Basico";
   "Entradas_Stopper" AT %E42.0 : "UDT_Entradas_Stopper";
   "Salidas_Basico" AT %A1.0 : "UDT_Salidas_Basico";
   "Salidas_APP" AT %A0.0 : "UDT_Salidas_APP";
   "Entradas_RFID" AT %E10.0 : "UDT_Entradas_RFID";
   "Salidas_RFID" AT %A10.0 : "UDT_Salidas_RFID";
END_VAR

VAR_GLOBAL CONSTANT   // PLC tag table "Tabla de variables estándar"
   "Ninguno" : Pip := 65535;
   "Actualización automática" : Pip := 0;
   "MIPP 1" : Pip := 1;
   "MIPP 2" : Pip := 2;
   "MIPP 3" : Pip := 3;
   "MIPP 4" : Pip := 4;
   "MIPP 5" : Pip := 5;
   "MIPP 6" : Pip := 6;
   "MIPP 7" : Pip := 7;
   "MIPP 8" : Pip := 8;
   "MIPP 9" : Pip := 9;
   "MIPP 10" : Pip := 10;
   "MIPP 11" : Pip := 11;
   "MIPP 12" : Pip := 12;
   "MIPP 13" : Pip := 13;
   "MIPP 14" : Pip := 14;
   "MIPP 15" : Pip := 15;
   "MIPP 16" : Pip := 16;
   "MIPP 17" : Pip := 17;
   "MIPP 18" : Pip := 18;
   "MIPP 19" : Pip := 19;
   "MIPP 20" : Pip := 20;
   "MIPP 21" : Pip := 21;
   "MIPP 22" : Pip := 22;
   "MIPP 23" : Pip := 23;
   "MIPP 24" : Pip := 24;
   "MIPP 25" : Pip := 25;
   "MIPP 26" : Pip := 26;
   "MIPP 27" : Pip := 27;
   "MIPP 28" : Pip := 28;
   "MIPP 29" : Pip := 29;
   "MIPP 30" : Pip := 30;
   "MIPP 31" : Pip := 31;
   "MIPP OB Servo" : Pip := 32768;
   "Local~MC" : Hw_SubModule := 51;
   "Local~Common" : Hw_SubModule := 50;
   "Local~Device" : Hw_Device := 32;
   "Local~Configuration" : Hw_SubModule := 33;
   "Local~Exec" : Hw_SubModule := 52;
   "Local" : Hw_SubModule := 49;
   "Local~FExec" : Hw_SubModule := 55;
   "Local~Interfaz_PROFINET_1" : Hw_Interface := 64;
   "Local~Interfaz_PROFINET_1~Puerto_3" : Hw_Interface := 67;
   "Local~Interfaz_PROFINET_1~Port_1" : Hw_Interface := 65;
   "Local~Interfaz_PROFINET_1~Port_2" : Hw_Interface := 66;
   "Local~DI_8x24VDC_HF_1" : Hw_SubModule := 257;
   "Local~DI_8x24VDC_HF_2" : Hw_SubModule := 258;
   "Local~DQ_8x24VDC_0_5A_HF_1" : Hw_SubModule := 259;
   "Local~DQ_8x24VDC_0_5A_HF_2" : Hw_SubModule := 260;
   "Local~CM_4xIO-Link_1" : Hw_SubModule := 261;
   "OB_Main" : OB_PCYCLE := 1;
   "Local~Módulo_servidor_1" : Hw_SubModule := 262;
END_VAR

// ===== library: MasterCopy "Est_FB_App_Plantilla" =====

FUNCTION_BLOCK "Est_FB_App_Plantilla"   // FB6, SCL
{ S7_Optimized_Access := 'TRUE' }
VERSION : 0.1
   VAR_INPUT
      Entradas_app : "UDT_Entradas_APP";   // UDT propio de la estacion: sensores de la aplicacion
      App_inicio : Bool;   // la estacion pide empezar (palet leido y en posicion)
      Emergencia : Bool;
      Rearme : Bool;   // flanco del boton de rearme
   END_VAR
   VAR_OUTPUT
      App_en_reposo : Bool;   // la aplicacion esta lista para recibir un palet
      App_terminada : Bool;   // la aplicacion ha acabado; la estacion escribe el tag
      App_alarma : Bool;   // parpadeo de alarma en el piloto q2 (opcional)
      App_rearme_requerido : Bool;   // enciende la luz de rearme (opcional)
      Inhibir_cinta : Bool;   // TRUE = la cinta no debe moverse (por ejemplo, eje fuera de reposo)
   END_VAR
   VAR_IN_OUT
      Salidas_app : "UDT_Salidas_APP";   // UDT propio de la estacion: actuadores de la aplicacion
      Imagen_palet : Array[0..27] of Byte;   // bloque del tag RFID: lee y escribe aqui, solo en tus bytes
   END_VAR
   VAR
      Etapa_app : Int;   // Bytes del tag que usa ESTA estacion. Ver Mapa_RFID_CPLab.xlsx. Tienen que estar dentro de Mascara_lectura / Mascara_escritura de Main.
   END_VAR
   VAR CONSTANT
      IDX_EJEMPLO_LEER : Int := 5;
      IDX_EJEMPLO_ESCRIBIR : Int := 4;
   END_VAR
BEGIN

   // Salidas a su valor seguro en cada ciclo; cada etapa activa las que necesite
   #App_en_reposo := FALSE;
   #App_terminada := FALSE;
   #App_alarma := FALSE;
   #Inhibir_cinta := FALSE;

   CASE #Etapa_app OF
       0:  // REPOSO
           // TODO: condicion real de reposo de tu estacion (sensores en posicion inicial)
           #App_en_reposo := TRUE;
           IF #App_inicio AND #App_en_reposo THEN
               // Ejemplo de lectura de un byte del tag:
               //   IF #Imagen_palet[#IDX_EJEMPLO_LEER] = 1 THEN ...
               #Etapa_app := 10;
           END_IF;

       10: // TRABAJO
           // TODO: secuencia de tu estacion. Activa aqui tus Salidas_app.
           // Ejemplo de escritura de un byte del tag (solo si esta en Mascara_escritura):
           //   #Imagen_palet[#IDX_EJEMPLO_ESCRIBIR] := #Imagen_palet[#IDX_EJEMPLO_ESCRIBIR] OR 16#01;
           #Etapa_app := 20;

       20: // FIN: se mantiene hasta que la estacion baja App_inicio
           #App_terminada := TRUE;
           IF NOT #App_inicio THEN
               #Etapa_app := 0;
           END_IF;

       ELSE
           #Etapa_app := 0;
   END_CASE;

   // Emergencia: todo a seguro y vuelta a reposo
   IF #Emergencia THEN
       #Etapa_app := 0;
       // TODO: pon a FALSE todas tus Salidas_app
   END_IF;
   // TODO si tu estacion necesita rearme propio: App_rearme_requerido := TRUE hasta que llegue #Rearme
END_FUNCTION_BLOCK